// TIA Portal V21 export
FUNCTION_BLOCK "FB_Mixed"   // FB9, LAD
TITLE = KOP-Baustein mit SCL-Netzwerk / LAD block with an SCL network
{ S7_Optimized_Access := 'TRUE' }
// stored: MemoryReserve 100, SetENOAutomatically false
   VAR_INPUT
      Start : Bool;   // Startbefehl / Start command
      RawValue : Int;   // Rohwert / Raw value
   END_VAR
   VAR_OUTPUT
      Running : Bool;   // Läuft / Running
      Scaled : Real;   // Skalierter Wert / Scaled value
      AboveLimit : Bool;   // Läuft und über dem Grenzwert / Running and above the limit
   END_VAR
   VAR
      Factor : Real := 2.5;   // Skalierungsfaktor / Scaling factor
      Limit : Real := 100.0;   // Grenzwert / Limit
      IsAbove : Bool;   // Skalierter Wert über dem Grenzwert / Scaled value above the limit
   END_VAR
BEGIN

REGION Network 1: KOP-Netzwerk vor dem SCL-Netzwerk / LAD network before the SCL network
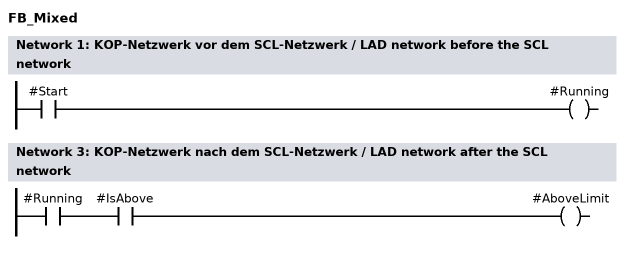
   RUNG wire#powerrail
      Contact( #Start )
      Coil( #Running )
   END_RUNG
   // the same network as SCL:
   #Running := #Start;
END_REGION

REGION Network 2 (SCL): SCL-Netzwerk im KOP-Baustein / SCL network inside the LAD block

       // Scale the raw value and compare it with the limit
       #Scaled := INT_TO_REAL(#RawValue) * #Factor;
       #IsAbove := #Scaled > #Limit;
END_REGION

REGION Network 3: KOP-Netzwerk nach dem SCL-Netzwerk / LAD network after the SCL network
   RUNG wire#powerrail
      Contact( #Running )
      Contact( #IsAbove )
      Coil( #AboveLimit )
   END_RUNG
   // the same network as SCL:
   #AboveLimit := #Running AND #IsAbove;
END_REGION
END_FUNCTION_BLOCK
